PROGRAM main
  VAR
    MARCHA AT %IX0.0  : BOOL; (* S1, pulsador NA *)
    PARADA AT %IX0.1  : BOOL; (* S2, pulsador NC *)
    TERMICO AT %IX0.2 : BOOL; (* F1, térmico NC *)
    KM1 AT %QX0.0     : BOOL; (* contactor del motor *)
    H1 AT %QX0.1      : BOOL; (* piloto de falla *)
    H2 AT %QX0.2      : BOOL; (* piloto de marcha *)
    FALLA             : BOOL; (* falla del térmico memorizada *)
    RS_KM1            : RS;
    SR_FALLA          : SR;
  END_VAR
  VAR  (* added by the conversion: wires and edge detectors of the diagram *)
    _NOT4_OUT : BOOL;
    _NOT6_OUT : BOOL;
    _OR3_OUT : BOOL;
  END_VAR

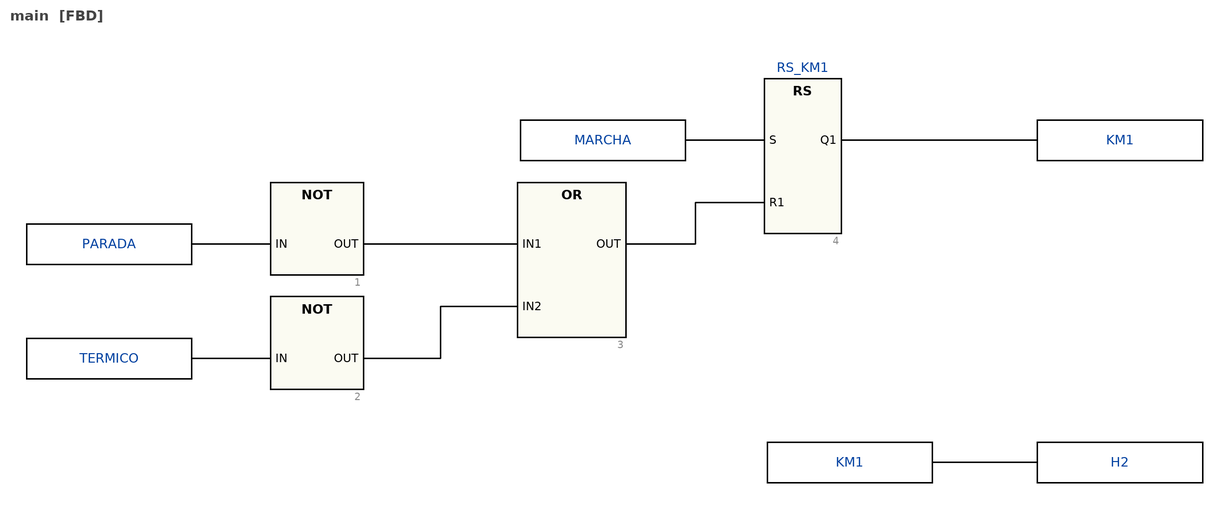
(* FBD diagram, written out as Structured Text *)
_NOT4_OUT := NOT PARADA;
_NOT6_OUT := NOT TERMICO;
_OR3_OUT := _NOT4_OUT OR _NOT6_OUT;
RS_KM1(S := MARCHA, R1 := _OR3_OUT);
KM1 := RS_KM1.Q1;
H2 := KM1;
END_PROGRAM
